# EPICS substitutions: xrmIocApp/Db/permit_AI_16CH.substitutions
file "permit_AI.template"
{
	pattern {CH, ADDR}
        {ALL, 0}
	{01, 1}
	{02, 2}
	{03, 3}
	{04, 4}
	{05, 5}
	{06, 6}
	{07, 7}
	{08, 8}
	{09, 9}
	{10,10}
	{11,11}
	{12,12}
	{13,13}
	{14,14}
	{15,15}
	{16,16}
}
